// TIA Portal project "Week1_1" (V20)

(* hardware
DEVICE "S7-1200 station_1"  S7-1200 Station
   slot 0: "Rack_0"  S7-1200 Rack  Rack  V1.0
   slot 1: "PLC_1"  CPU 1214C AC/DC/Rly  6ES7 214-1BG40-0XB0  V4.6
DEVICE "PC-System_1"  SIMATIC PC station
   slot 0: "SIMATIC PC station"  Rail  SIMATIC PC-Station  V1.0
      slot 125: "Stationmanager"  Station_Manager  V6.0.4
   slot 1: "HMI_RT_1"  WinCC RT Advanced  6AV2 104-0xxxx-xxxx  17.0.0.0
      slot 33792: "Computer interface"  Host interface
   slot 2: "IE general_1"  IE General  IE_CP  V8.2.0
      slot 1: "PROFINET interface"  IEGeneral.Interface.8.2.0
*)

// ===== PLC "PLC_1"  CPU 1214C AC/DC/Rly =====

VAR_GLOBAL   // PLC tag table "Default tag table"
   "System_Byte" AT %MB1 : Byte;
   "FirstScan" AT %M1.0 : Bool;
   "DiagStatusUpdate" AT %M1.1 : Bool;
   "AlwaysTRUE" AT %M1.2 : Bool;
   "AlwaysFALSE" AT %M1.3 : Bool;
   "Clock_Byte" AT %MB0 : Byte;
   "Clock_10Hz" AT %M0.0 : Bool;
   "Clock_5Hz" AT %M0.1 : Bool;
   "Clock_2.5Hz" AT %M0.2 : Bool;
   "Clock_2Hz" AT %M0.3 : Bool;
   "Clock_1.25Hz" AT %M0.4 : Bool;
   "Clock_1Hz" AT %M0.5 : Bool;
   "Clock_0.625Hz" AT %M0.6 : Bool;
   "Clock_0.5Hz" AT %M0.7 : Bool;
   "SW1" AT %M2.0 : Bool;
   "SW2" AT %M2.1 : Bool;
   "SW3" AT %M2.2 : Bool;
   "SW4" AT %M2.3 : Bool;
   "LED1" AT %M3.0 : Bool;
   "LED2" AT %M3.1 : Bool;
   "LED3" AT %M3.2 : Bool;
   "LED4" AT %M3.3 : Bool;
END_VAR

DATA_BLOCK "DB_Array"   // DB1
{ S7_Optimized_Access := 'TRUE' }
VERSION : 0.1
   VAR
      Count : Int;
      QR_Code : Array[1..10] of Struct
         QR_Source : String;
         Count : Int;
      END_STRUCT;
      QR_Read : String;
      Order : Int;
      Ready : Bool;
   END_VAR
BEGIN
END_DATA_BLOCK

ORGANIZATION_BLOCK "Main"   // OB1, LAD, ProgramCycle
TITLE = "Main Program Sweep (Cycle)"
{ S7_Optimized_Access := 'TRUE' }
VERSION : 0.1
   VAR_INPUT
      Initial_Call : Bool;   // Initial call of this OB
      Remanence : Bool;   // =True, if remanent data are available
   END_VAR
   VAR_TEMP
      i : Int;
   END_VAR
BEGIN

REGION Network 1
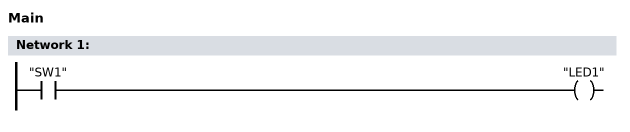
   RUNG wire#powerrail
      Contact( "SW1" )
      Coil( "LED1" )
   END_RUNG
   // the same network as SCL:
   "LED1" := "SW1";
END_REGION

REGION Network 2 (SCL)
   // อ่านคิวอาร์
   IF "DB_Array".Ready THEN
       FOR #i := 1 TO 10 DO
           IF "DB_Array".QR_Read = "DB_Array".QR_Code[#i].QR_Source THEN
               "DB_Array".QR_Code[#i].Count := "DB_Array".QR_Code[#i].Count + "DB_Array".Order;
               "DB_Array".Ready := 0;
               RETURN;

           END_IF;
       END_FOR;

       FOR #i := 1 TO 10 DO
           IF "DB_Array".QR_Code[#i]."QR_Source" =  '' THEN
               "DB_Array".QR_Code[#i].QR_Source := "DB_Array".QR_Read;
               "DB_Array".QR_Code[#i].Count := "DB_Array".QR_Code[#i].Count + "DB_Array".Order;
               EXIT;
           END_IF;
       END_FOR;
       "DB_Array".Ready := 0;
   END_IF;
END_REGION
END_ORGANIZATION_BLOCK

(* ===== HMI "HMI_RT_1" =====
system functions are stored by id; their names below are inferred from use
connection "HMI_Connection_1": ETHERNET, S7_1200_OMS

HMI tags "Default tag table"
   "LED1" : Bool = PLC LED1 AT %M3.0, 1 s
   "SW1" : Bool = PLC SW1 AT %M2.0, 1 s
   "DB_Array_QR_Read" : String[254] = PLC DB_Array.QR_Read, 1 s
   "DB_Array_Order" : Int = PLC DB_Array.Order, 1 s
   "DB_Array_Ready" : Bool = PLC DB_Array.Ready, 1 s
   "DB_Array_QR_Code{0}_QR_Source" : String[254] = PLC DB_Array.QR_Code[1].QR_Source, 1 s
   "DB_Array_QR_Code{0}_Count" : Int = PLC DB_Array.QR_Code[1].Count, 1 s
   "DB_Array_QR_Code{1}_QR_Source" : String[254] = PLC DB_Array.QR_Code[1].QR_Source, 1 s
   "DB_Array_QR_Code{1}_Count" : Int = PLC DB_Array.QR_Code[1].Count, 1 s
   "DB_Array_QR_Code{2}_QR_Source" : String[254] = PLC DB_Array.QR_Code[2].QR_Source, 1 s
   "DB_Array_QR_Code{2}_Count" : Int = PLC DB_Array.QR_Code[2].Count, 1 s
   "DB_Array_QR_Code{3}_QR_Source" : String[254] = PLC DB_Array.QR_Code[3].QR_Source, 1 s
   "DB_Array_QR_Code{3}_Count" : Int = PLC DB_Array.QR_Code[3].Count, 1 s
   "DB_Array_QR_Code{4}_QR_Source" : String[254] = PLC DB_Array.QR_Code[4].QR_Source, 1 s
   "DB_Array_QR_Code{4}_Count" : Int = PLC DB_Array.QR_Code[4].Count, 1 s
   "DB_Array_QR_Code{5}_Count" : Int = PLC DB_Array.QR_Code[5].Count, 1 s
   "DB_Array_QR_Code{5}_QR_Source" : String[254] = PLC DB_Array.QR_Code[5].QR_Source, 1 s
   "DB_Array_QR_Code{6}_QR_Source" : String[254] = PLC DB_Array.QR_Code[6].QR_Source, 1 s
   "DB_Array_QR_Code{7}_QR_Source" : String[254] = PLC DB_Array.QR_Code[7].QR_Source, 1 s
   "DB_Array_QR_Code{8}_QR_Source" : String[254] = PLC DB_Array.QR_Code[8].QR_Source, 1 s
   "DB_Array_QR_Code{9}_QR_Source" : String[254] = PLC DB_Array.QR_Code[9].QR_Source, 1 s
   "DB_Array_QR_Code{10}_QR_Source" : String[254] = PLC DB_Array.QR_Code[10].QR_Source, 1 s
   "DB_Array_QR_Code{6}_Count" : Int = PLC DB_Array.QR_Code[6].Count, 1 s
   "DB_Array_QR_Code{7}_Count" : Int = PLC DB_Array.QR_Code[7].Count, 1 s
   "DB_Array_QR_Code{8}_Count" : Int = PLC DB_Array.QR_Code[8].Count, 1 s
   "DB_Array_QR_Code{9}_Count" : Int = PLC DB_Array.QR_Code[9].Count, 1 s
   "DB_Array_QR_Code{10}_Count" : Int = PLC DB_Array.QR_Code[10].Count, 1 s

screen "Screen_1" 1024x768
   TextField "Text field_1" at 41,37 size 134x29; Text 'Automation'
   Circle "Circle_1" at 69,85 size 75x75
      Appearance <- "LED1"
   Button "Button_2" at 171,176 size 96x32; TextOff 'SW1'
      on Press: SetBit("SW1")
      on Release: ResetBit("SW1")
   Button "Button_1" at 13,176 size 135x32; TextOff 'SW1 InvertBit'
      on Click: InvertBit("SW1")
   TextField "Text field_3" at 385,151 size 43x22; Text 'สินค้า'
   IOField "I/O field_1" at 384,181 size 167x32; FormatPattern ????????????????????????????????????????????????????????????????????????????????
      ProcessValue <- "DB_Array_QR_Code{1}_QR_Source"
   IOField "I/O field_2" at 624,178 size 96x32; FormatPattern s99999
      ProcessValue <- "DB_Array_QR_Code{1}_Count"
   TextField "Text field_4" at 617,153 size 50x22; Text 'จำนวน'
   TextField "Text field_2" at 363,46 size 127x22; Text 'ช่องรับ QR-CODE'
   IOField "I/O field_3" at 368,72 size 149x32; FormatPattern ??????????????????????????????????????????????????
      ProcessValue <- "DB_Array_QR_Read"
   TextField "Text field_5" at 554,46 size 50x22; Text 'จำนวน'
   IOField "I/O field_4" at 543,71 size 109x32; FormatPattern s999999
      ProcessValue <- "DB_Array_Order"
   Button "Button_3" at 686,68 size 96x32; TextOff 'ยืนยัน'
      on Click: SetBit("DB_Array_Ready")
   IOField "I/O field_5" at 385,219 size 167x32; FormatPattern ????????????????????????????????????????????????????????????????????????????????
      ProcessValue <- "DB_Array_QR_Code{2}_QR_Source"
   IOField "I/O field_6" at 385,255 size 167x32; FormatPattern ????????????????????????????????????????????????????????????????????????????????
      ProcessValue <- "DB_Array_QR_Code{3}_QR_Source"
   IOField "I/O field_7" at 385,292 size 167x32; FormatPattern ????????????????????????????????????????????????????????????????????????????????
      ProcessValue <- "DB_Array_QR_Code{4}_QR_Source"
   IOField "I/O field_8" at 385,330 size 167x32; FormatPattern ????????????????????????????????????????????????????????????????????????????????
      ProcessValue <- "DB_Array_QR_Code{5}_QR_Source"
   IOField "I/O field_9" at 385,366 size 167x32; FormatPattern ????????????????????????????????????????????????????????????????????????????????
      ProcessValue <- "DB_Array_QR_Code{6}_QR_Source"
   IOField "I/O field_10" at 384,401 size 167x32; FormatPattern ????????????????????????????????????????????????????????????????????????????????
      ProcessValue <- "DB_Array_QR_Code{7}_QR_Source"
   IOField "I/O field_11" at 384,441 size 167x32; FormatPattern ????????????????????????????????????????????????????????????????????????????????
      ProcessValue <- "DB_Array_QR_Code{8}_QR_Source"
   IOField "I/O field_12" at 384,478 size 167x32; FormatPattern ????????????????????????????????????????????????????????????????????????????????
      ProcessValue <- "DB_Array_QR_Code{9}_QR_Source"
   IOField "I/O field_13" at 384,514 size 167x32; FormatPattern ????????????????????????????????????????????????????????????????????????????????
      ProcessValue <- "DB_Array_QR_Code{10}_QR_Source"
   IOField "I/O field_14" at 623,218 size 96x32; FormatPattern s99999
      ProcessValue <- "DB_Array_QR_Code{2}_Count"
   IOField "I/O field_15" at 623,255 size 96x32; FormatPattern s99999
      ProcessValue <- "DB_Array_QR_Code{3}_Count"
   IOField "I/O field_16" at 622,330 size 96x32; FormatPattern s99999
      ProcessValue <- "DB_Array_QR_Code{5}_Count"
   IOField "I/O field_17" at 623,293 size 96x32; FormatPattern s99999
      ProcessValue <- "DB_Array_QR_Code{4}_Count"
   IOField "I/O field_18" at 623,368 size 96x32; FormatPattern s99999
      ProcessValue <- "DB_Array_QR_Code{6}_Count"
   IOField "I/O field_19" at 623,402 size 96x32; FormatPattern s99999
      ProcessValue <- "DB_Array_QR_Code{7}_Count"
   IOField "I/O field_20" at 623,440 size 96x32; FormatPattern s99999
      ProcessValue <- "DB_Array_QR_Code{8}_Count"
   IOField "I/O field_21" at 622,476 size 96x32; FormatPattern s99999
      ProcessValue <- "DB_Array_QR_Code{9}_Count"
   IOField "I/O field_22" at 622,515 size 96x32; FormatPattern s99999
      ProcessValue <- "DB_Array_QR_Code{10}_Count"
*)